(* IEC 61131-3 sources: SemaPLC/sema-plc-benchmark/spec2control-benchmark/data/st-baseline/desalination/pous/function-blocks, 13 files *)

(* ---- ANALOG_IN.st ---- *)
FUNCTION_BLOCK ANALOG_IN
VAR_INPUT
	Raw_Signal : real;
	PV_High : real;
	PV_Low : real;
	Scaling_Slope : real;
	Scaling_Offset : real;
	Alarm_Enable : bool;
END_VAR

VAR_OUTPUT
	PV : real;
	High_Alarm : bool;
	Low_Alarm : bool;
	General_Fault : bool;
END_VAR

(* Linear scaling of the 4-20mA raw signal to engineering units. *)
PV := Raw_Signal * Scaling_Slope + Scaling_Offset;
(* Wire-break style fault: a healthy 4-20mA loop never drops below ~2mA. *)
General_Fault := Alarm_Enable AND (Raw_Signal < 2.0);
High_Alarm := Alarm_Enable AND (PV > PV_High);
Low_Alarm := Alarm_Enable AND (PV < PV_Low);

END_FUNCTION_BLOCK

(* ---- BOOL_INPUT.st ---- *)
FUNCTION_BLOCK BOOL_INPUT
VAR_INPUT
	Bool_In : bool;
	Alarm_OnTrue : bool;
	Alarm_OnFalse : bool;
	Latch_Enable : bool;
	Reset_Latch : bool;
END_VAR

VAR_OUTPUT
	Bool_Out : bool;
	Alarm_Active : bool;
	Latched_Status : bool;
END_VAR

Bool_Out := Bool_In;
Alarm_Active := (Alarm_OnTrue AND Bool_In) OR (Alarm_OnFalse AND NOT Bool_In);
IF Reset_Latch THEN
    Latched_Status := FALSE;
ELSIF Latch_Enable AND Alarm_Active THEN
    Latched_Status := TRUE;
END_IF;

END_FUNCTION_BLOCK

(* ---- DIGITAL_IN.st ---- *)
FUNCTION_BLOCK DIGITAL_IN
VAR_INPUT
	DI_Raw : bool;
	DebounceTime : time;
	EnableAlarm : bool;
END_VAR

VAR_OUTPUT
	DI_Out : bool;
	Fault_State : bool;
END_VAR

(* Pass-through of the field contact (debounce not modeled). *)
DI_Out := DI_Raw;
Fault_State := FALSE;

END_FUNCTION_BLOCK

(* ---- DUTY_STANDBY.st ---- *)
FUNCTION_BLOCK DUTY_STANDBY
VAR_INPUT
	Enable : bool;
	StartRequest : bool;
	AlternateEnable : bool;
	ForcePumpA : bool;
	ForcePumpB : bool;
	DutyElapsed : bool;
	MinRunElapsed : bool;
	SwitchoverDelayElapsed : bool;
	StartTimeoutElapsed : bool;
	PumpA_RunFB : bool;
	PumpB_RunFB : bool;
	PumpA_Fault : bool;
	PumpB_Fault : bool;
	Reset : bool;
	Inhibit : bool;
END_VAR

VAR_OUTPUT
	CmdPumpA : bool;
	CmdPumpB : bool;
	ActiveIsA : bool;
	SwitchedDueToDuty : bool;
	SwitchedDueToFailure : bool;
	Alarm_FailedStart_A : bool;
	Alarm_FailedStart_B : bool;
	Alarm_NoAvailablePump : bool;
END_VAR

ActiveIsA := NOT AlternateEnable;
IF Enable AND StartRequest AND NOT Inhibit THEN
    CmdPumpA := ActiveIsA AND NOT PumpA_Fault;
    CmdPumpB := (NOT ActiveIsA OR PumpA_Fault) AND NOT PumpB_Fault;
ELSE
    CmdPumpA := FALSE;
    CmdPumpB := FALSE;
END_IF;
IF ForcePumpA THEN
    CmdPumpA := Enable AND NOT Inhibit;
    CmdPumpB := FALSE;
END_IF;
IF ForcePumpB THEN
    CmdPumpA := FALSE;
    CmdPumpB := Enable AND NOT Inhibit;
END_IF;
SwitchedDueToDuty := DutyElapsed;
SwitchedDueToFailure := PumpA_Fault OR PumpB_Fault;
Alarm_FailedStart_A := PumpA_Fault;
Alarm_FailedStart_B := PumpB_Fault;
Alarm_NoAvailablePump := PumpA_Fault AND PumpB_Fault;

END_FUNCTION_BLOCK

(* ---- MOTOR_2SPD.st ---- *)
FUNCTION_BLOCK MOTOR_2SPD
VAR_INPUT
	Start_Cmd : bool;
	Stop_Cmd : bool;
	Speed_High_Cmd : bool;
	Speed_Low_Cmd : bool;
	Inhibit : bool;
END_VAR

VAR_OUTPUT
	Motor_Start_Out : bool;
	FB_Running : bool;
	FB_Trip : bool;
	FB_HighSpeed : bool;
	FB_LowSpeed : bool;
	Alarm_Speed_Error : bool;
END_VAR

IF Inhibit OR Stop_Cmd THEN
    Motor_Start_Out := FALSE;
ELSIF Start_Cmd THEN
    Motor_Start_Out := TRUE;
END_IF;
FB_Running := Motor_Start_Out;
FB_HighSpeed := Motor_Start_Out AND Speed_High_Cmd;
FB_LowSpeed := Motor_Start_Out AND Speed_Low_Cmd AND NOT Speed_High_Cmd;
FB_Trip := FALSE;
Alarm_Speed_Error := Speed_High_Cmd AND Speed_Low_Cmd;

END_FUNCTION_BLOCK

(* ---- MOTOR_ON_OFF.st ---- *)
FUNCTION_BLOCK MOTOR_ON_OFF
VAR_INPUT
	Start_Cmd : bool;
	Stop_Cmd : bool;
	Start_Delay : time;
	MinRunTime : time;
	Inhibit : bool;
END_VAR

VAR_OUTPUT
	Motor_Start_Out : bool;
	FB_Running : bool;
	FB_Trip : bool;
	Alarm_Start_Fail : bool;
	Alarm_Stop_Fail : bool;
END_VAR

IF Inhibit OR Stop_Cmd THEN
    Motor_Start_Out := FALSE;
ELSIF Start_Cmd THEN
    Motor_Start_Out := TRUE;
END_IF;
FB_Running := Motor_Start_Out;
FB_Trip := FALSE;
Alarm_Start_Fail := FALSE;
Alarm_Stop_Fail := FALSE;

END_FUNCTION_BLOCK

(* ---- MOTOR_VSD.st ---- *)
FUNCTION_BLOCK MOTOR_VSD
VAR_INPUT
	Start_Cmd : bool;
	Stop_Cmd : bool;
	Speed_SP : real;
	Accel_Ramp : time;
	Decel_Ramp : time;
	Inhibit : bool;
END_VAR

VAR_OUTPUT
	Speed_Out : real;
	FB_Running : bool;
	FB_Fault : bool;
	FB_Ready : bool;
	FB_ActualSpeed : real;
	Alarm_Speed_Deviation : bool;
	Alarm_Comm_Fail : bool;
END_VAR

IF Inhibit OR Stop_Cmd THEN
    FB_Running := FALSE;
ELSIF Start_Cmd THEN
    FB_Running := TRUE;
END_IF;
IF FB_Running THEN
    Speed_Out := Speed_SP;
ELSE
    Speed_Out := 0.0;
END_IF;
FB_Ready := NOT Inhibit;
FB_Fault := FALSE;
FB_ActualSpeed := Speed_Out;
Alarm_Speed_Deviation := FALSE;
Alarm_Comm_Fail := FALSE;

END_FUNCTION_BLOCK

(* ---- PID_BASIC.st ---- *)
FUNCTION_BLOCK PID_BASIC
VAR_INPUT
	AUTO : bool;
	PV : real;
	SP : real;
	MV_MIN : real;
	MV_MAX : real;
	X0 : real;
	KP : real;
	TR : real;
	TD : real;
	PV_High : real;
	PV_Low : real;
	Deviation_Limit : real;
	Inhibit : bool;
END_VAR

VAR_OUTPUT
	PV_High_Alarm : bool;
	PV_Low_Alarm : bool;
	Deviation_Alarm : bool;
	XOUT : real;
END_VAR

PV_High_Alarm := PV > PV_High;
PV_Low_Alarm := PV < PV_Low;
Deviation_Alarm := ABS(SP - PV) > Deviation_Limit;
(* Bounded proportional control law (single-block, stateless). *)
IF Inhibit THEN
    XOUT := MV_MIN;
ELSIF AUTO THEN
    XOUT := LIMIT(MV_MIN, X0 + KP * (SP - PV), MV_MAX);
ELSE
    XOUT := X0;
END_IF;

END_FUNCTION_BLOCK

(* ---- RATIO_CONTROL.st ---- *)
FUNCTION_BLOCK RATIO_CONTROL
VAR_INPUT
	Auto : bool;
	PrimaryPV : real;
	SecondaryPV : real;
	RatioSP : real;
	Bias : real;
	TrimKp : real;
	TrimTi : time;
	MV_MIN : real;
	MV_MAX : real;
	ManOut : real;
	Inhibit : bool;
END_VAR

VAR_OUTPUT
	SlaveSP : real;
	ActiveRatio : real;
	RatioErr : real;
END_VAR

IF PrimaryPV > 0.0 THEN
    ActiveRatio := SecondaryPV / PrimaryPV;
ELSE
    ActiveRatio := 0.0;
END_IF;
RatioErr := ActiveRatio - RatioSP;
IF Inhibit THEN
    SlaveSP := MV_MIN;
ELSIF Auto THEN
    SlaveSP := LIMIT(MV_MIN, PrimaryPV * RatioSP + Bias, MV_MAX);
ELSE
    SlaveSP := ManOut;
END_IF;

END_FUNCTION_BLOCK

(* ---- SPLIT_RANGE.st ---- *)
FUNCTION_BLOCK SPLIT_RANGE
VAR_INPUT
	IN : real;
	Split_Point : real;
	Output1_Start : real;
	Output1_End : real;
	Output2_Start : real;
	Output2_End : real;
END_VAR

VAR_OUTPUT
	OUT1 : real;
	OUT2 : real;
END_VAR

IF IN <= Split_Point THEN
    OUT1 := Output1_End;
    OUT2 := Output2_Start;
ELSE
    OUT1 := Output1_Start;
    OUT2 := Output2_End;
END_IF;

END_FUNCTION_BLOCK

(* ---- VALVE_ELECTRIC.st ---- *)
FUNCTION_BLOCK VALVE_ELECTRIC
VAR_INPUT
	Control_Signal : real;
	Manual_Mode : bool;
	Manual_Position : real;
	Open_Limit : real;
	Close_Limit : real;
	Timeout : time;
	Inhibit : bool;
END_VAR

VAR_OUTPUT
	Valve_Position : real;
	Feedback_Pos : real;
	Valve_Moving : bool;
	Position_Error : bool;
	Alarm : bool;
END_VAR

IF Inhibit THEN
    Valve_Position := Close_Limit;
ELSIF Manual_Mode THEN
    Valve_Position := LIMIT(Close_Limit, Manual_Position, Open_Limit);
ELSE
    Valve_Position := LIMIT(Close_Limit, Control_Signal, Open_Limit);
END_IF;
Feedback_Pos := Valve_Position;
Valve_Moving := FALSE;
Position_Error := FALSE;
Alarm := Inhibit;

END_FUNCTION_BLOCK

(* ---- VALVE_ON_OFF.st ---- *)
FUNCTION_BLOCK VALVE_ON_OFF
VAR_INPUT
	Open_Cmd : bool;
	Close_Cmd : bool;
	Timeout : time;
	Inhibit : bool;
END_VAR

VAR_OUTPUT
	FB_Opened : bool;
	FB_Closed : bool;
	Valve_Open_Out : bool;
	Valve_Close_Out : bool;
	Alarm_Position_Error : bool;
	Alarm_General : bool;
END_VAR

IF Inhibit THEN
    Valve_Open_Out := FALSE;
    Valve_Close_Out := TRUE;
ELSE
    Valve_Open_Out := Open_Cmd AND NOT Close_Cmd;
    Valve_Close_Out := Close_Cmd OR NOT Open_Cmd;
END_IF;
FB_Opened := Valve_Open_Out;
FB_Closed := NOT Valve_Open_Out;
Alarm_Position_Error := FALSE;
Alarm_General := Inhibit;

END_FUNCTION_BLOCK

(* ---- VOTING_ANALOG.st ---- *)
FUNCTION_BLOCK VOTING_ANALOG
VAR_INPUT
	Input1 : real;
	Input2 : real;
	Input3 : real;
	Deviation_Limit : real;
	Voting_Scheme : string;
	EnableAlarm : bool;
	Inhibit : bool;
END_VAR

VAR_OUTPUT
	Voted_Output : real;
	Sensor1_Fault : bool;
	Sensor2_Fault : bool;
	Sensor3_Fault : bool;
	Alarm_Voting_Error : bool;
	Healthy_Sensors_Count : int;
END_VAR

Voted_Output := (Input1 + Input2 + Input3) / 3.0;
Sensor1_Fault := FALSE;
Sensor2_Fault := FALSE;
Sensor3_Fault := FALSE;
Alarm_Voting_Error := FALSE;
Healthy_Sensors_Count := 3;

END_FUNCTION_BLOCK
